(*
SPDX-FileCopyrightText: c 2026 Oleksandr Tiutyk <trofimich@gmail.com>
SPDX-License-Identifier: MIT
License: https://opensource.org/license/mit
*)

(*!
<summary>Checks clearing a full inline index and refilling with distinct values.</summary>
<description>
Owns a fixed-capacity set and copied values at a stable address. Run from one task.
Teardown clears surviving entries before publication.
</description>
*)

{attribute 'no_assign'}
{attribute 'no_explicit_call' := 'do not call this function block directly'}
FUNCTION_BLOCK StaticUniqueDataSetClearTest EXTENDS TOF_Testing.SingleCycleTest
VAR_STAT
	{attribute 'hide'}
	_ClassName : STRING := __POUNAME();
END_VAR
VAR
	_Set : TOF_Collections.UniqueDataSet<7>(valueValidator := 0, valueEqualityComparer := 0);
END_VAR

(*!
<summary>Checks clearing a full inline index and refilling with distinct values.</summary>
*)
METHOD PROTECTED ExecuteTest
VAR
	values : ARRAY [0..6] OF STRING :=
		['String0', 'String1', 'String2', 'String3', 'String4', 'String5', 'String6'];
	i : DINT;
	replacementValues : ARRAY [0..6] OF INT := [11, 12, 13, 14, 15, 16, 17];
END_VAR
FOR i := 6 TO 0 BY -1 DO
	_Set.SetCopy(value := values[i]);
END_FOR

Assert.ThatBool(
	actual := _Set.Full AND_THEN _Set.Length = 7,
	message := "The clear fixture must start full"
).IsTrue();

_Set.Clear();

Assert.ThatBool(
	actual := _Set.Empty AND_THEN _Set.Length = 0 AND_THEN NOT _Set.Full,
	message := "Clearing a full set must make every slot available"
).IsTrue();

Assert.ThatDInt(
	actual := _Set.Capacity,
	message := "Clearing must preserve inline capacity"
).ToBe(expected := DINT#7);

FOR i := 0 TO 6 DO
	Assert.ThatBool(
		actual := _Set.Contains(value := values[i]),
		message := TOF_Core.WideStrings.Concat255("Clear must hide the old value at offset ", TO_WSTRING(i))
	).IsFalse();
END_FOR

FOR i := 0 TO 6 DO
	_Set.SetCopy(value := replacementValues[i]);
END_FOR

Assert.ThatBool(
	actual := _Set.Full AND_THEN _Set.Length = 7,
	message := "Refilling must reuse all seven slots"
).IsTrue();

FOR i := 0 TO 6 DO
	Assert.ThatBool(
		actual := _Set.Contains(value := replacementValues[i]),
		message := TOF_Core.WideStrings.Concat255("Refill must index value ", TO_WSTRING(replacementValues[i]))
	).IsTrue();
END_FOR
END_METHOD

(*!
<summary>Clears the fixture before the runner publishes the result.</summary>
<description>
Also runs after an unexpected exception interrupts the case.
</description>
*)
METHOD PROTECTED AfterTest
_Set.Clear();
END_METHOD

//! <summary>Borrows the concrete class name. Callers must not modify it.</summary>
{attribute 'monitoring' := 'call'}
PROPERTY ClassName : REFERENCE TO STRING
GET
ClassName REF= _ClassName;
END_GET
END_PROPERTY

//! <summary>Borrows the compiler-initialized namespace name. Callers must not modify it.</summary>
{attribute 'monitoring' := 'call'}
PROPERTY NamespaceName : REFERENCE TO STRING
GET
NamespaceName REF= CurrentNamespace.Name;
END_GET
END_PROPERTY

//! <summary>Reports the concrete instance size in bytes.</summary>
{attribute 'monitoring' := 'call'}
PROPERTY SelfSize : ULINT
GET
SelfSize := XSIZEOF(THIS^);
END_GET
END_PROPERTY

END_FUNCTION_BLOCK

(* stored: Version 1.1.0.1
   POU StaticUniqueDataSetClearTest: Id {e6ef3022-5dc9-4c79-b0a6-b5287548122e}, SpecialFunc None
   Method ExecuteTest: Id {c056d05c-4835-49fe-9711-23f84aebd11d}
   Method AfterTest: Id {c41766a4-84f4-4fb3-8832-5e854726f698}
   Property ClassName: Id {4a35889c-7fc0-4218-b286-95d4f08fbd76}
   Get Get: Id {e83ad39f-e278-40ad-9ccf-4b2464d8267c}
   Property NamespaceName: Id {9626d720-766e-4928-8d46-d88ace1390da}
   Get Get: Id {4691424a-0ffa-40a2-9968-8538c51bf56a}
   Property SelfSize: Id {1d0aba78-2e53-4512-b72c-f8572251da94}
   Get Get: Id {e2e0b742-a622-4b9b-8211-7bc0c8d10609} *)
